Fanuc KAREL source: kt00441.KL

-- PROVISIONAL review KL for V770-1; original PC SHA256 ee557a8c3c6043d54073ffd9a71396f0e99098a1d868abc3b822a7b49cd67b7c
-- Incomplete behavior may be omitted. Consult companion uncertainty JSON. Do not deploy.
PROGRAM KT00441
%NOLOCKGROUP
VAR
  R1 : REAL
  I2 : INTEGER
  OUT : BOOLEAN
BEGIN
  -- UNRESOLVED_PC offsets 5-16; opcodes 2E,23
  -- UNRESOLVED_PC offsets 21-32; opcodes 2E,23
  -- UNRESOLVED_PC offsets 37-57; opcodes 21,21,64,72,23
  -- UNRESOLVED_PC offsets 62-66; opcodes 7F
END KT00441
